(* IEC 61131-3 sources: codesys-framework/txt/application/WeVe General (library)/CsvFileLogger/FB_CsvFileLogger/Properties, 3 files *)

(* ---- Count.prop.st ---- *)
// Aantal regels dat nog in de buffer wacht.
PROPERTY Count : INT
// --- BEGIN IMPLEMENTATION ---

// ----------- GET -----------
VAR
END_VAR

// -- BEGIN IMPLEMENTATION GET --
Count := _iCount;

(* ---- Error.prop.st ---- *)
// TRUE zolang het bestand niet geschreven kan worden (de logger probeert om de tRetry opnieuw).
PROPERTY Error : BOOL
// --- BEGIN IMPLEMENTATION ---

// ----------- GET -----------
VAR
END_VAR

// -- BEGIN IMPLEMENTATION GET --
Error := _xError;

(* ---- Overflow.prop.st ---- *)
// Totaal aantal regels dat verloren ging omdat de buffer vol was.
PROPERTY Overflow : UDINT
// --- BEGIN IMPLEMENTATION ---

// ----------- GET -----------
VAR
END_VAR

// -- BEGIN IMPLEMENTATION GET --
Overflow := _udiOverflow;
